# EPICS substitutions: iocs/motor/pi-ioc/db/PI_C663.substitutions
# PI_C663.substitutions, as C's iocPI has for its other controllers,
# on this IOC's axes, P and C from st.cmd; the values are the motor
# record this IOC had before.
#
# PI C-663: one motor record for the controller's single axis, DTYP "PIC663"
# with OUT #C$(C) S0, as the C-862 it clones.
#
# The C-663 works in raw controller counts (MA/MR/TP are integer counts, no
# separate EGU scaling in the driver), so MRES = 1 and EGU = counts.
file "$(MOTOR)/db/motor.db"
{
pattern
{M,       DTYP,      S,  DESC,  EGU,     DIR,  VELO,  VBAS,  ACCL,  BDST,  BVEL,  BACC,  MRES,  PREC,  DHLM,     DLLM,      INIT}
{"c663",  "PIC663",  0,  "",    counts,  Pos,  1000,  0,     0.2,   0,     0,     .5,    1,     0,     1000000,  -1000000,  ""}
}
